// TIA Portal project "EXO1" (V16)

(* hardware
DEVICE "Station S7300/ET200M_1"  S7-300 station
   slot 0: "Châssis_0"  Rail  6ES7 390-1***0-0AA0
   slot 1: "PS 307 10A_1"  PS 307 10A  6ES7 307-1KA02-0AA0
   slot 2: "PLC_1"  CPU 314  6ES7 314-1AG13-0AB0  V2.6
      slot 0: "Interface MPI_1"  X1
   slot 4: "DI 16x24VDC_1"  DI16 x 24VDC, interrupt  6ES7 321-7BH01-0AB0
   slot 5: "DO 8x24VDC/0.5A_1"  DO8 x 24VDC / 0.5A  6ES7 322-8BF00-0AB0
*)

// ===== PLC "PLC_1"  CPU 314 =====

VAR_GLOBAL   // PLC tag table "Table de variables standard"
   "BP_MARCHE" AT %I0.0 : Bool;
   "BP_ARRET" AT %I0.1 : Bool;
   "lampe1" AT %Q0.2 : Bool;
   "lampe2" AT %Q0.3 : Bool;
   "moteur" AT %Q0.4 : Bool;
END_VAR

ORGANIZATION_BLOCK "Main"   // OB1, LAD
TITLE = "Main Program Sweep (Cycle)"
{ S7_Optimized_Access := 'FALSE' }
VERSION : 0.1
   VAR_TEMP
      OB1_EV_CLASS : Byte;   // Bits 0-3 = 1 (Coming event), Bits 4-7 = 1 (Event class 1)
      OB1_SCAN_1 : Byte;   // 1 (Cold restart scan 1 of OB 1), 3 (Scan 2-n of OB 1)
      OB1_PRIORITY : Byte;   // Priority of OB Execution
      OB1_OB_NUMBR : Byte;   // 1 (Organization block 1, OB1)
      OB1_RESERVED_1 : Byte;   // Reserved for system
      OB1_RESERVED_2 : Byte;   // Reserved for system
      OB1_PREV_CYCLE : Int;   // Cycle time of previous OB1 scan (milliseconds)
      OB1_MIN_CYCLE : Int;   // Minimum cycle time of OB1 (milliseconds)
      OB1_MAX_CYCLE : Int;   // Maximum cycle time of OB1 (milliseconds)
      OB1_DATE_TIME : Date_And_Time;   // Date and time OB1 started
   END_VAR
BEGIN

REGION Network 1
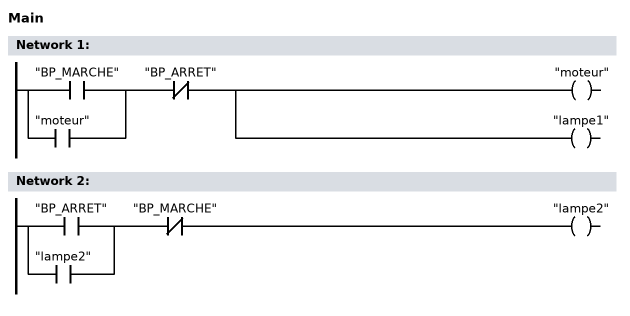
   RUNG wire#powerrail
      Contact( "BP_MARCHE" )
      wire#w1
      I_Contact( "BP_ARRET" )
      wire#w2
      Coil( "moteur" )
   END_RUNG
   RUNG wire#powerrail
      Contact( "moteur" )
   END_RUNG wire#w1
   RUNG wire#w2
      Coil( "lampe1" )
   END_RUNG
   // the same network as SCL:
   "moteur" := ("BP_MARCHE" OR "moteur") AND NOT "BP_ARRET";
   "lampe1" := "moteur";
END_REGION

REGION Network 2
   RUNG wire#powerrail
      Contact( "BP_ARRET" )
      wire#w1
      I_Contact( "BP_MARCHE" )
      Coil( "lampe2" )
   END_RUNG
   RUNG wire#powerrail
      Contact( "lampe2" )
   END_RUNG wire#w1
   // the same network as SCL:
   "lampe2" := ("BP_ARRET" OR "lampe2") AND NOT "BP_MARCHE";
END_REGION
END_ORGANIZATION_BLOCK